SUBAPPLICATION Uebung_006g_AX (* SR-Flip-Flop via INIT_ON_OFF, ausgeloest von 2x E_TRIG (EInitOn/EInitOff Broadcast auf unverbundene Events) *)
  (* Standard: 61499-2; Description: Copyright (c) 2026 Meisterschulen am Ostbahnhof This program and the accompanying materials are made available under the terms of the Eclipse Public License 2.0 which is available at https://www.eclipse.org/legal/epl-2.0/ SPDX-License-Identifier: EPL-2.0 *)
  (* Version 1.0, 2026-10-11, Franz Höpfinger, Meisterschulen am Ostbahnhof, initial API and implementation and/or initial documentation *)
  PACKAGE Uebungen;
  IMPORT logiBUS::io::DI::logiBUS_DI::Input_I1;
  IMPORT logiBUS::io::DI::logiBUS_DI::Input_I2;
  IMPORT logiBUS::io::DI::logiBUS_DI_Events::BUTTON_SINGLE_CLICK;
  IMPORT logiBUS::io::DQ::logiBUS_DO::Output_Q1;
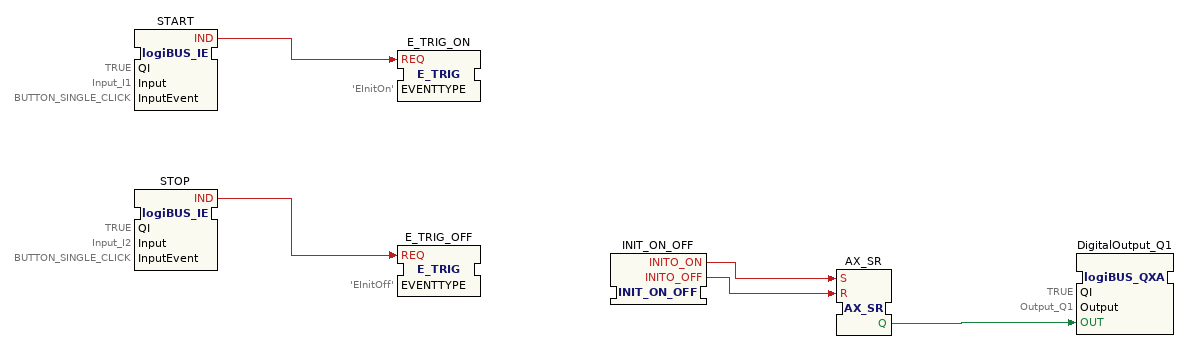
  (* INIT_ON und INIT_OFF bleiben unverbunden: E_TRIG broadcastet sein EVENTTYPE auf ALLE unverbundenen Events dieses Typs im Netzwerk - daher reagiert hier nur der passende Kanal (EInitOn bzw. EInitOff). *)
  FBS
    DigitalOutput_Q1 : logiBUS::io::DQ::logiBUS_QXA(QI := TRUE, Output := Output_Q1);
    START : logiBUS::io::DI::logiBUS_IE(QI := TRUE, Input := Input_I1, InputEvent := BUTTON_SINGLE_CLICK);
    STOP : logiBUS::io::DI::logiBUS_IE(QI := TRUE, Input := Input_I2, InputEvent := BUTTON_SINGLE_CLICK);
    E_TRIG_ON : iec61499::events::E_TRIG(EVENTTYPE := 'EInitOn');
    E_TRIG_OFF : iec61499::events::E_TRIG(EVENTTYPE := 'EInitOff');
    INIT_ON_OFF : events::init::INIT_ON_OFF;
    AX_SR : adapter::events::unidirectional::AX_SR;
  END_FBS
  EVENT_CONNECTIONS
    START.IND TO E_TRIG_ON.REQ;
    STOP.IND TO E_TRIG_OFF.REQ;
    INIT_ON_OFF.INITO_ON TO AX_SR.S;
    INIT_ON_OFF.INITO_OFF TO AX_SR.R;
  END_CONNECTIONS
  ADAPTER_CONNECTIONS
    AX_SR.Q TO DigitalOutput_Q1.OUT;
  END_CONNECTIONS
END_SUBAPPLICATION
